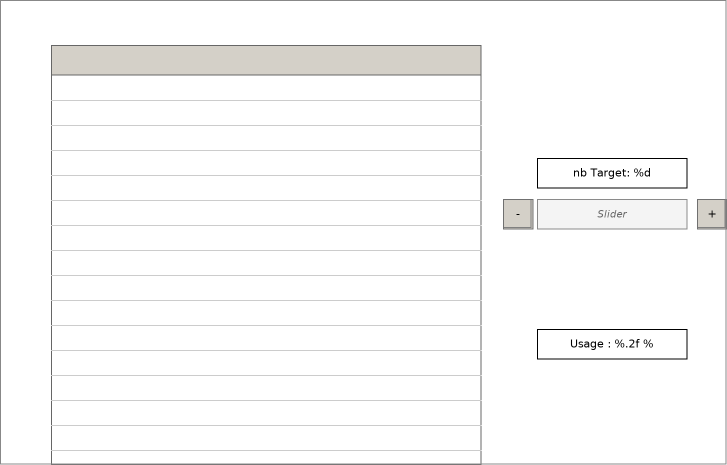
VISUALIZATION Visualization  // 727x465
    Table (51,45 430x420), data array: multiInstances.aFB
        p1128707560: multiInstances.cMaxInstances
        p3854506369: multiInstances.aFB[INDEX]^.nCounts
        p1014161805: MULTIINSTANCES.cMaxInstances - 1 + INT#1
    Rectangle (537,158 150x30), "nb Target: %d", text variable: multiInstances.nTarget
        OnMouseClick: write the text variable via Default, min 1, max multiInstances.cMaxInstances
    Rectangle (537,329 150x30), "Usage : %.2f %", text variable: multiInstances.nUsage
    Slider (537,199 150x30), variable: multiInstances.nTarget, scale 1..100
    Button (697,199 30x30), "+"
        OnMouseClick: toggle multiInstances.bInc
    Button (503,199 30x30), "-"
        OnMouseClick: toggle multiInstances.bDec
END_VISUALIZATION

(* stored: Version 1.1.0.1, ProductVersion 3.1.4026.21
   Visu Visualization: Id {b1108311-c32d-4723-94af-8d1a050141ea} *)
